(* IEC 61131-3 sources: llm-plc-st-eval/codesys/dobles/B6, 7 files *)

(* ---- 01_CorrectaInicioOFF.st ---- *)
(* DOBLE DE PRUEBA B6/CorrectaInicioOFF - NO ES CORPUS. Esperado: veredicto 1 *)
FUNCTION_BLOCK FB_Baliza
VAR_INPUT
    alarma : BOOL;
END_VAR
VAR_OUTPUT
    lampara : BOOL;
END_VAR
VAR
    t1 : TON;
    t2 : TON;
    prevAlarma : BOOL;
END_VAR
IF NOT alarma THEN
    lampara := FALSE;
    t1(IN := FALSE, PT := T#1S);
    t2(IN := FALSE, PT := T#1S);
    prevAlarma := FALSE;
ELSE
    prevAlarma := TRUE;
    IF lampara THEN
        t1(IN := FALSE, PT := T#1S);
        t2(IN := TRUE, PT := T#1S);
        IF t2.Q THEN
            lampara := FALSE;
        END_IF
    ELSE
        t2(IN := FALSE, PT := T#1S);
        t1(IN := TRUE, PT := T#1S);
        IF t1.Q THEN
            lampara := TRUE;
        END_IF
    END_IF
END_IF
END_FUNCTION_BLOCK

(* ---- 02_CorrectaInicioON.st ---- *)
(* DOBLE DE PRUEBA B6/CorrectaInicioON - NO ES CORPUS. Esperado: veredicto 1 *)
FUNCTION_BLOCK FB_Baliza
VAR_INPUT
    alarma : BOOL;
END_VAR
VAR_OUTPUT
    lampara : BOOL;
END_VAR
VAR
    t1 : TON;
    t2 : TON;
    prevAlarma : BOOL;
END_VAR
IF NOT alarma THEN
    lampara := FALSE;
    t1(IN := FALSE, PT := T#1S);
    t2(IN := FALSE, PT := T#1S);
    prevAlarma := FALSE;
ELSE
    IF NOT prevAlarma THEN
        lampara := TRUE;             (* enciende en el flanco de alarma *)
    END_IF
    prevAlarma := TRUE;
    IF lampara THEN
        t1(IN := FALSE, PT := T#1S);
        t2(IN := TRUE, PT := T#1S);
        IF t2.Q THEN
            lampara := FALSE;
        END_IF
    ELSE
        t2(IN := FALSE, PT := T#1S);
        t1(IN := TRUE, PT := T#1S);
        IF t1.Q THEN
            lampara := TRUE;
        END_IF
    END_IF
END_IF
END_FUNCTION_BLOCK

(* ---- 03_Periodo1500.st ---- *)
(* DOBLE DE PRUEBA B6/Periodo1500 - NO ES CORPUS. Esperado: veredicto 2, falla en el paso 1 *)
FUNCTION_BLOCK FB_Baliza
VAR_INPUT
    alarma : BOOL;
END_VAR
VAR_OUTPUT
    lampara : BOOL;
END_VAR
VAR
    t1 : TON;
    t2 : TON;
    prevAlarma : BOOL;
END_VAR
IF NOT alarma THEN
    lampara := FALSE;
    t1(IN := FALSE, PT := T#1500MS);
    t2(IN := FALSE, PT := T#1500MS);
    prevAlarma := FALSE;
ELSE
    IF NOT prevAlarma THEN
        lampara := TRUE;             (* enciende en el flanco de alarma *)
    END_IF
    prevAlarma := TRUE;
    IF lampara THEN
        t1(IN := FALSE, PT := T#1500MS);
        t2(IN := TRUE, PT := T#1500MS);
        IF t2.Q THEN
            lampara := FALSE;
        END_IF
    ELSE
        t2(IN := FALSE, PT := T#1500MS);
        t1(IN := TRUE, PT := T#1500MS);
        IF t1.Q THEN
            lampara := TRUE;
        END_IF
    END_IF
END_IF
END_FUNCTION_BLOCK

(* ---- 04_Periodo500.st ---- *)
(* DOBLE DE PRUEBA B6/Periodo500 - NO ES CORPUS. Esperado: veredicto 2, falla en el paso 1 *)
FUNCTION_BLOCK FB_Baliza
VAR_INPUT
    alarma : BOOL;
END_VAR
VAR_OUTPUT
    lampara : BOOL;
END_VAR
VAR
    t1 : TON;
    t2 : TON;
    prevAlarma : BOOL;
END_VAR
IF NOT alarma THEN
    lampara := FALSE;
    t1(IN := FALSE, PT := T#500MS);
    t2(IN := FALSE, PT := T#500MS);
    prevAlarma := FALSE;
ELSE
    IF NOT prevAlarma THEN
        lampara := TRUE;             (* enciende en el flanco de alarma *)
    END_IF
    prevAlarma := TRUE;
    IF lampara THEN
        t1(IN := FALSE, PT := T#500MS);
        t2(IN := TRUE, PT := T#500MS);
        IF t2.Q THEN
            lampara := FALSE;
        END_IF
    ELSE
        t2(IN := FALSE, PT := T#500MS);
        t1(IN := TRUE, PT := T#500MS);
        IF t1.Q THEN
            lampara := TRUE;
        END_IF
    END_IF
END_IF
END_FUNCTION_BLOCK

(* ---- 05_Asimetrico.st ---- *)
(* DOBLE DE PRUEBA B6/Asimetrico - NO ES CORPUS. Esperado: veredicto 2, falla en el paso 1 *)
FUNCTION_BLOCK FB_Baliza
VAR_INPUT
    alarma : BOOL;
END_VAR
VAR_OUTPUT
    lampara : BOOL;
END_VAR
VAR
    t1 : TON;
    t2 : TON;
    prevAlarma : BOOL;
END_VAR
IF NOT alarma THEN
    lampara := FALSE;
    t1(IN := FALSE, PT := T#2S);
    t2(IN := FALSE, PT := T#1S);
    prevAlarma := FALSE;
ELSE
    IF NOT prevAlarma THEN
        lampara := TRUE;             (* enciende en el flanco de alarma *)
    END_IF
    prevAlarma := TRUE;
    IF lampara THEN
        t1(IN := FALSE, PT := T#2S);
        t2(IN := TRUE, PT := T#1S);
        IF t2.Q THEN
            lampara := FALSE;
        END_IF
    ELSE
        t2(IN := FALSE, PT := T#1S);
        t1(IN := TRUE, PT := T#2S);
        IF t1.Q THEN
            lampara := TRUE;
        END_IF
    END_IF
END_IF
END_FUNCTION_BLOCK

(* ---- 06_SiempreEncendida.st ---- *)
(* DOBLE DE PRUEBA B6/SiempreEncendida - NO ES CORPUS. Esperado: veredicto 2, falla en el paso 1 *)
FUNCTION_BLOCK FB_Baliza
VAR_INPUT
    alarma : BOOL;
END_VAR
VAR_OUTPUT
    lampara : BOOL;
END_VAR
VAR
    nada : BOOL;
END_VAR
lampara := alarma;
END_FUNCTION_BLOCK

(* ---- 07_NoApagaSinAlarma.st ---- *)
(* DOBLE DE PRUEBA B6/NoApagaSinAlarma - NO ES CORPUS. Esperado: veredicto 2, falla en el paso 2 *)
FUNCTION_BLOCK FB_Baliza
VAR_INPUT
    alarma : BOOL;
END_VAR
VAR_OUTPUT
    lampara : BOOL;
END_VAR
VAR
    t1 : TON;
    t2 : TON;
    prevAlarma : BOOL;
    visto : BOOL;
    alarmaEf : BOOL;
END_VAR
IF alarma THEN
    visto := TRUE;
END_IF
alarmaEf := visto OR alarma;
IF NOT alarmaEf THEN
    lampara := FALSE;
    t1(IN := FALSE, PT := T#1S);
    t2(IN := FALSE, PT := T#1S);
    prevAlarma := FALSE;
ELSE
    IF NOT prevAlarma THEN
        lampara := TRUE;             (* enciende en el flanco de alarma *)
    END_IF
    prevAlarma := TRUE;
    IF lampara THEN
        t1(IN := FALSE, PT := T#1S);
        t2(IN := TRUE, PT := T#1S);
        IF t2.Q THEN
            lampara := FALSE;
        END_IF
    ELSE
        t2(IN := FALSE, PT := T#1S);
        t1(IN := TRUE, PT := T#1S);
        IF t1.Q THEN
            lampara := TRUE;
        END_IF
    END_IF
END_IF
END_FUNCTION_BLOCK
